(*
SPDX-FileCopyrightText: © 2026 Oleksandr Tiutyk <trofimich@gmail.com>
SPDX-License-Identifier: MIT
License: https://opensource.org/license/mit
*)

(*!
<summary>Defines relational and equality comparison operators for workflow conditions.</summary>
*)

{attribute 'qualified_only'}
{attribute 'strict'}
{attribute 'to_string'}
TYPE COMPARISON_OPERATOR :
(
	EQUAL := 0,
	NOT_EQUAL := 1,
	LESS_THAN := 2,
	LESS_THAN_OR_EQUAL := 3,
	GREATER_THAN := 4,
	GREATER_THAN_OR_EQUAL := 5
) BYTE;
END_TYPE

(* stored: Version 1.1.0.1
   DUT COMPARISON_OPERATOR: Id {6915700c-027c-4794-9bf1-95f9336a12c2} *)
